(*
SPDX-FileCopyrightText: c 2026 Oleksandr Tiutyk <trofimich@gmail.com>
SPDX-License-Identifier: MIT
License: https://opensource.org/license/mit
*)

(*!
<summary>Checks removal of all matches while preserving the order of survivors.</summary>
<description>
Borrows a group-owned list reserved for this case. Use from one task at a stable address.
Teardown clears the list before publication.
</description>
*)

{attribute 'no_assign'}
{attribute 'no_explicit_call' := 'do not call this function block directly'}
FUNCTION_BLOCK ListRemoveMatchedTest EXTENDS TOF_Testing.SingleCycleTest
VAR_STAT
	{attribute 'hide'}
	_ClassName : STRING := __POUNAME();
END_VAR
VAR
	_List : TOF_Collections.IList;
	_Predicate : ListStringPredicate;
END_VAR

(*!
<summary>Clears the fixture before the runner publishes the result.</summary>
<description>
Also runs after an unexpected exception interrupts the case.
</description>
*)
METHOD PROTECTED AfterTest
_List.Clear();
END_METHOD

//! <summary>Borrows the concrete class name. Callers must not modify it.</summary>
{attribute 'monitoring' := 'call'}
PROPERTY ClassName : REFERENCE TO STRING
GET
ClassName REF= _ClassName;
END_GET
END_PROPERTY

(*!
<summary>Checks removal of all matches while preserving the order of survivors.</summary>
*)
METHOD PROTECTED ExecuteTest
VAR
	values : ARRAY [0..5] OF STRING := ['String0', 'String1', 'String2', 'String3', 'String4', 'String5'];
	expected : ARRAY [0..5] OF STRING := ['String0', 'String1', 'String3', 'String4', 'String5', 'String3'];
	i : DINT;
END_VAR
_List.AppendCopy(value := values[0]);
_List.AppendCopy(value := values[1]);
_List.AppendCopy(value := values[2]);
_List.AppendCopy(value := values[3]);
_List.AppendCopy(value := values[4]);
_List.AppendCopy(value := values[5]);
_List.AppendCopy(value := values[2]);
_List.AppendCopy(value := values[3]);

_Predicate.Expected := 'String2';
_List.RemoveMatched(predicate := _Predicate);

Assert.ThatDInt(
	actual := _List.Length,
	message := "Unexpected sequence after RemoveMatched length"
).ToBe(expected := DINT#6);

FOR i := 0 TO 5 DO
	Assert.ThatString(
		actual := _List.Get(index := i).AsString255(),
		message := TOF_Core.WideStrings.Concat255("Unexpected sequence after RemoveMatched at index ", TO_WSTRING(i))
	).ToBe(expected := expected[i]);
END_FOR
END_METHOD

(*!
<summary>Binds the list fixture for this case.</summary>
<description>
Stores a borrowed interface without invoking the fixture. The owning group keeps it alive and
reserves it for this case. TestElement initializes the name and parent.
</description>
<param name="name">Display name of this case.</param>
<param name="parent">Group that owns this case.</param>
<param name="list">Required live list reserved for this case.</param>
*)
METHOD FB_init : BOOL
VAR_INPUT
	bInitRetains: BOOL; // TRUE: the retain variables are initialized (reset warm / reset cold)
	bInCopyCode: BOOL; // TRUE: the instance will be copied to the copy code afterward (online change)
	name : WSTRING;
	parent : TOF_Testing.ITestElement;
	list : TOF_Collections.IList;
END_VAR
_List := list;
FB_init := TRUE;
END_METHOD

//! <summary>Borrows the compiler-initialized namespace name. Callers must not modify it.</summary>
{attribute 'monitoring' := 'call'}
PROPERTY NamespaceName : REFERENCE TO STRING
GET
NamespaceName REF= CurrentNamespace.Name;
END_GET
END_PROPERTY

//! <summary>Reports the concrete instance size in bytes.</summary>
{attribute 'monitoring' := 'call'}
PROPERTY SelfSize : ULINT
GET
SelfSize := XSIZEOF(THIS^);
END_GET
END_PROPERTY

END_FUNCTION_BLOCK

(* stored: Version 1.1.0.1, ProductVersion 3.1.4026.21
   POU ListRemoveMatchedTest: Id {50db1e6c-87b1-4ae3-921f-0eb309c43ee7}, SpecialFunc None
   Method AfterTest: Id {594dfe6d-185f-462f-b55a-486e60fd2a08}
   Property ClassName: Id {5876a3bd-69da-4a95-8d6e-553b3dfa1fde}
   Get Get: Id {835b8abe-849c-411e-b0f6-b7659257d1e3}
   Method ExecuteTest: Id {88070a78-7720-4cab-8435-c008e40b32d2}
   Method FB_init: Id {1ce24023-47d5-42d9-ae74-bc8b1fe0c18a}
   Property NamespaceName: Id {716c67c8-7255-4bce-86e3-ece140e3eb87}
   Get Get: Id {7d07c533-043a-469b-a15b-7c4582f68144}
   Property SelfSize: Id {68cfa4fc-6611-43ff-9305-e0f90f944f6f}
   Get Get: Id {3909eac3-4720-4027-adef-11ac2a45b1c8} *)
